Fanuc KAREL source: KA00175.KL

PROGRAM KA00175
%NOLOCKGROUP
VAR
  SRC: ARRAY[4] OF STRING[20]
  DST: ARRAY[4] OF STRING[20]
BEGIN
  DST = SRC
END KA00175
